Staubli VAL3: getPath.pgx

program getPath(string x_sHmiName, string& x_sHmiPath)
begin
  x_sHmiPath=libPath()+"/interface/"+x_sHmiName
end
